// TIA Portal V19 export
TYPE "SKID_VFD"
   STRUCT
      START_CMD : Bool;
      FAULT_RESET : Bool;
      RUN_FBK : Bool;
      TRIP_FBK : Bool;
      LOCAL_REMOTE : Bool;
      SPEED_REF : Real;
      SPEED_ACT : Real;
   END_STRUCT;
END_TYPE
